# EPICS autosave request: vme_iocs/iocbio4/iocBoot/ioc18IDd/auto_positions.req
$(P)m1.DVAL
$(P)m2.DVAL
$(P)m3.DVAL
$(P)m4.DVAL
$(P)m5.DVAL
$(P)m6.DVAL
$(P)m7.DVAL
$(P)m8.DVAL
$(P)m9.DVAL
$(P)m10.DVAL
$(P)m11.DVAL
$(P)m12.DVAL
$(P)m13.DVAL
$(P)m14.DVAL
$(P)m15.DVAL
$(P)m16.DVAL
